(* IEC 61131-3 sources: kns-port-domestic/upstream/plc-process-lib/src/DUTs/Pid, 6 files *)

(* ---- E_PidAction.dut.st ---- *)
// Назначение: направление действия ПИД-регулятора.
// Автор:      kr0nsch
// Версия:     0.1.0
// Документ:   docs/fb/FB_PID.md
{attribute 'qualified_only'}
{attribute 'strict'}
TYPE E_PidAction :
(
    Reverse := 0,   // обратное: PV растёт — выход падает (e = SP − PV); нагрев, подача
    Direct  := 1    // прямое: PV растёт — выход растёт (e = PV − SP); уровень → скорость откачки
) INT;
END_TYPE

(* ---- E_PidAlarm.dut.st ---- *)
// Назначение: индексы слотов тревог ПИД-регулятора. Нестрогое перечисление: им
//             индексируются массивы.
// Автор:      kr0nsch
// Версия:     0.1.0
// Документ:   docs/fb/FB_PID.md
{attribute 'qualified_only'}
TYPE E_PidAlarm :
(
    PvInvalid := 0   // PV недостоверна в Auto
) UINT;
END_TYPE

(* ---- E_PidPvFailAction.dut.st ---- *)
// Назначение: реакция ПИД-регулятора в Auto на недостоверную PV.
// Автор:      kr0nsch
// Версия:     0.1.0
// Документ:   docs/fb/FB_PID.md
{attribute 'qualified_only'}
{attribute 'strict'}
TYPE E_PidPvFailAction :
(
    Hold         := 0,   // удерживать выход; когда PV снова годна — продолжить без рывка
    SafeOut      := 1,   // выход := rSafeOut_pct; возврат без рывка
    ShedToManual := 2    // перейти в Manual с текущим выходом; в Auto возвращает оператор
) INT;
END_TYPE

(* ---- ST_PidCfg.dut.st ---- *)
// Назначение: параметры ПИД-регулятора (Persistent Variables приложения,
//             VAR_IN_OUT CONSTANT stCfg). Значения по умолчанию проходят CheckConfig.
//             Тип лежит в Persistent Variables приложения и заморожен в пределах 1.x (A-13).
// Автор:      kr0nsch
// Версия:     0.1.0
// Документ:   docs/fb/FB_PID.md
{attribute 'qualified_only'}
TYPE ST_PidCfg :
STRUCT
    eAction        : E_PidAction := E_PidAction.Reverse;
    rKp            : REAL := 1.0;     // %/% (выход в % на % диапазона PV); знак — только через eAction
    rTi_s          : REAL := 30.0;    // 0 — без И (интегратор = смещение, задаётся предустановкой)
    rTd_s          : REAL := 0.0;     // 0 — без Д
    rDFilterN      : REAL := 10.0;    // фильтр Д: Tf = Td / N
    rTt_s          : REAL := 0.0;     // постоянная слежения anti-windup; 0 — авто
    rPvMin_eu      : REAL := 0.0;     // диапазон PV для нормировки (как у датчика)
    rPvMax_eu      : REAL := 100.0;
    rSpMin_eu      : REAL := 0.0;     // пределы задания
    rSpMax_eu      : REAL := 100.0;
    rSpRate_ups    : REAL := 0.0;     // рампа задания, инж. ед./с; 0 — нет
    rOutMin_pct    : REAL := 0.0;     // пределы выхода
    rOutMax_pct    : REAL := 100.0;
    rOutRate_pctps : REAL := 0.0;     // ограничение скорости выхода, %/с; 0 — нет
    rDeadband_pct  : REAL := 0.0;     // зона нечувствительности по ошибке, % диапазона PV
    tSample        : TIME := T#0S;    // период расчёта; T#0S — каждый вызов
    tDtMax         : TIME := T#2S;    // больший шаг — разрыв (стоп ПЛК, отладка): шаг пропускается
    ePvFailAction  : E_PidPvFailAction := E_PidPvFailAction.Hold;
    rSafeOut_pct   : REAL := 0.0;     // выход при ePvFailAction = SafeOut
    xSpTrackPv     : BOOL := FALSE;   // в Manual задание следует за PV
    xUseOutAct     : BOOL := FALSE;   // обратный расчёт по rOutAct_pct (внешнее насыщение)
    udiAlarmIdBase : UDINT := 0;      // номер первой тревоги устройства (dev_no * 10)
    astAlarm       : ARRAY[0..GVL_Const.DEV_ALARMS_MAX - 1] OF ST_AlarmCfg := [
        (ePriority := E_AlarmPriority.Medium),    // 0 PvInvalid
        (ePriority := E_AlarmPriority.None), (ePriority := E_AlarmPriority.None),
        (ePriority := E_AlarmPriority.None), (ePriority := E_AlarmPriority.None),
        (ePriority := E_AlarmPriority.None), (ePriority := E_AlarmPriority.None),
        (ePriority := E_AlarmPriority.None)];
END_STRUCT
END_TYPE

(* ---- ST_PidCmd.dut.st ---- *)
// Назначение: команды HMI/SCADA ПИД-регулятора (GVL_Hmi приложения, VAR_IN_OUT stCmd).
// Автор:      kr0nsch
// Версия:     0.1.0
// Документ:   docs/fb/FB_PID.md
{attribute 'qualified_only'}
TYPE ST_PidCmd :
STRUCT
    stCommon       : ST_DeviceCmd;   // xSetAuto, xSetManual, xSetOos, xReset, xAck ...
    rSp_eu         : REAL;           // задание оператора; при xSpExt ФБ пишет сюда внешнее
    rManualOut_pct : REAL;           // выход в Manual, %; в Auto/Track/OOS ФБ пишет сюда текущий выход
END_STRUCT
END_TYPE

(* ---- ST_PidSts.dut.st ---- *)
// Назначение: состояние ПИД-регулятора для HMI/SCADA. 64 байта, 32 регистра Modbus:
//             только 16- и 32-битные поля без скрытого выравнивания.
// Автор:      kr0nsch
// Версия:     0.1.0
// Документ:   docs/fb/FB_PID.md
{attribute 'qualified_only'}
TYPE ST_PidSts :
STRUCT
    stCommon     : ST_DeviceSts;   // 0..27
    rSpTarget_eu : REAL;   // 28: задание после пределов, до рампы
    rSp_eu       : REAL;   // 32: действующее задание (после рампы)
    rPv_eu       : REAL;   // 36: регулируемая величина
    rErr_pct     : REAL;   // 40: ошибка, % диапазона PV, со знаком действия, после зоны нечувствительности
    rOut_pct     : REAL;   // 44: выход
    rP_pct       : REAL;   // 48: пропорциональная составляющая
    rI_pct       : REAL;   // 52: интегральная составляющая
    rD_pct       : REAL;   // 56: дифференциальная составляющая
    rDt_ms       : REAL;   // 60: последний шаг расчёта
END_STRUCT
END_TYPE
